(* IEC 61131-3 sources: openplc-editor-canopen/src/backend/shared/transpilers/st-transpiler/__tests__/fixtures/ld-relayout-corpus/ld-corpus-hard/expected-st, 5 files *)

(* ---- _project.st ---- *)
CONFIGURATION Config0

  RESOURCE Res0 ON PLC
    TASK task0(INTERVAL := T#20ms,PRIORITY := 1);
    PROGRAM instance0 WITH task0 : main;
  END_RESOURCE
END_CONFIGURATION

(* ---- Chains.st ---- *)
PROGRAM Chains
  VAR
    h07_start : BOOL;
    TON0 : TON;
    CTU0 : CTU;
    h07_done : BOOL;
    h07_reset : BOOL;
    h07_count : INT;
    h08_start : BOOL;
    TON1 : TON;
    TOF0 : TOF;
    CTU1 : CTU;
    h08_done : BOOL;
    h08_r1 : BOOL;
    h08_r2 : BOOL;
    h08_count : INT;
  END_VAR

  TON0(IN := h07_start, PT := T#1s);
  CTU0(CU := TON0.Q, R := h07_reset, PV := 4);
  h07_done := CTU0.Q;
  h07_count := CTU0.CV;
  TON1(IN := h08_start, PT := T#1s);
  TOF0(IN := TON1.Q, PT := T#2s);
  CTU1(CU := TOF0.Q, R := h08_r1 OR h08_r2, PV := 3);
  h08_done := CTU1.Q;
  h08_count := CTU1.CV;
END_PROGRAM

(* ---- Counters.st ---- *)
PROGRAM Counters
  VAR
    h01_a : BOOL;
    CTU0 : CTU;
    h01_q : BOOL;
    h01_b : BOOL;
    h01_c : BOOL;
    h01_d : BOOL;
    h01_cv : INT;
    h02_a : BOOL;
    CTUD0 : CTUD;
    h02_qu : BOOL;
    h02_b : BOOL;
    h02_c : BOOL;
    h02_d : BOOL;
    h02_e : BOOL;
    h02_g : BOOL;
    h02_f : BOOL;
    h02_h : BOOL;
    h02_i : BOOL;
    h02_k : BOOL;
    h02_j : BOOL;
    h02_qd : BOOL;
    h02_cv : INT;
    h03_a : BOOL;
    SR0 : SR;
    h03_q1 : BOOL;
    h03_c : BOOL;
    h03_b : BOOL;
    h03_d : BOOL;
    h03_e : BOOL;
    RS0 : RS;
    h03_q2 : BOOL;
    h03_f : BOOL;
    h03_h : BOOL;
    h03_g : BOOL;
    h04_e : BOOL;
    TON0 : TON;
    h04_q : BOOL;
    h04_a : BOOL;
    h04_b : BOOL;
    h04_c : BOOL;
    h04_d : BOOL;
    h04_et : TIME;
  END_VAR

  CTU0(CU := h01_b AND h01_a, R := h01_c OR h01_d, PV := 10);
  h01_q := CTU0.Q;
  h01_cv := CTU0.CV;
  CTUD0(CU := (h02_b OR h02_d AND h02_c) AND h02_a, CD := h02_g AND (h02_e OR h02_f), R := h02_h, LD := h02_k OR h02_j AND h02_i, PV := 30);
  h02_qu := CTUD0.QU;
  h02_qd := CTUD0.QD;
  h02_cv := CTUD0.CV;
  SR0(S1 := h03_c AND (h03_a OR h03_b), R := h03_d);
  h03_q1 := SR0.Q1;
  RS0(S := h03_e, R1 := h03_h OR h03_g AND h03_f);
  h03_q2 := RS0.Q1;
  TON0(IN := h04_e OR (h04_b OR h04_d AND h04_c) AND h04_a, PT := T#3s);
  h04_q := TON0.Q;
  h04_et := TON0.ET;
END_PROGRAM

(* ---- Mixed.st ---- *)
PROGRAM Mixed
  VAR
    h10_a : BOOL;
    CTU0 : CTU;
    h10_q : BOOL;
    h10_r1 : BOOL;
    h10_r2 : BOOL;
    h10_cv : INT;
    h10_b : BOOL;
    TON0 : TON;
    h10_k1 : BOOL;
    h10_k2 : BOOL;
    h10_k3 : BOOL;
    h10_e : BOOL;
    h10_s : BOOL;
    SR0 : SR;
    h10_q1 : BOOL;
    h10_rr : BOOL;
  END_VAR

  CTU0(CU := h10_a, R := h10_r1 OR h10_r2, PV := 2);
  h10_q := CTU0.Q;
  h10_cv := CTU0.CV;
  TON0(IN := h10_b OR h10_e, PT := T#1s);
  h10_k1 := TON0.Q;
  h10_k2 := TON0.Q;
  h10_k3 := TON0.Q;
  SR0(S1 := h10_s, R := h10_rr);
  h10_q1 := SR0.Q1;
END_PROGRAM

(* ---- Parallel.st ---- *)
PROGRAM Parallel
  VAR
    TON0 : TON;
    h05_out : BOOL;
    CTU0 : CTU;
    h05_a : BOOL;
    h05_b : BOOL;
    h05_r : BOOL;
    h06_en : BOOL;
    h06_y1 : BOOL;
    h06_y2 : BOOL;
    h06_y3 : BOOL;
    h06_y4 : BOOL;
    TON1 : TON;
    h06_a1 : BOOL;
    TOF0 : TOF;
    h06_b1 : BOOL;
    CTU1 : CTU;
    h06_c1 : BOOL;
    h06_r : BOOL;
    h06_cv : INT;
    h09_out : BOOL;
    TON2 : TON;
    TOF1 : TOF;
    h09_a : BOOL;
    h09_b : BOOL;
    h09_c : BOOL;
    h09_d : BOOL;
    _TMP_AND5437823_OUT : BOOL;
  END_VAR

  TON0(IN := h05_a, PT := T#1s);
  CTU0(CU := h05_b, R := h05_r, PV := 5);
  h05_out := CTU0.Q OR TON0.Q;
  TON1(IN := h06_a1 AND h06_en, PT := T#1s);
  h06_y1 := TON1.Q;
  TOF0(IN := h06_b1 AND h06_en, PT := T#2s);
  h06_y2 := TOF0.Q;
  CTU1(CU := h06_c1 AND h06_en, R := h06_r, PV := 7);
  h06_y3 := CTU1.Q;
  h06_cv := CTU1.CV;
  h06_y4 := h06_en;
  TON2(IN := h09_a, PT := T#1s);
  TOF1(IN := h09_b, PT := T#2s);
  _TMP_AND5437823_OUT := AND(TOF1.Q OR TON2.Q, h09_c OR h09_d);
  h09_out := _TMP_AND5437823_OUT;
END_PROGRAM
